(* IEC 61131-3 sources: sis-interlock-demo/src/POUs/Sis/F_VoteArchRequired, 2 files *)

(* ---- F_VoteArchRequired.decl.st ---- *)
// Назначение: требуемое число голосов M схемы голосования по таблице 5.1; 0 — для None,
//             ForcedTrip и значений вне перечисления.
// Автор:      kr0nsch
// Версия:     0.1.0
// Документ:   docs/DESIGN.md, раздел «5.10 Вспомогательные функции голосования»
// ВНИМАНИЕ:   код демонстрационный и не предназначен для систем безопасности. Реальная ПАЗ
//             требует определения SIL, сертифицированных аппаратных и программных средств
//             и валидации по ГОСТ Р МЭК 61511.
FUNCTION F_VoteArchRequired : UINT
VAR_INPUT
    eArch : E_VoteArch;   // схема голосования
END_VAR

(* ---- F_VoteArchRequired.impl.st ---- *)
CASE eArch OF
    E_VoteArch.Vote1oo1, E_VoteArch.Vote1oo2:
        F_VoteArchRequired := 1;
    E_VoteArch.Vote2oo2, E_VoteArch.Vote2oo3:
        F_VoteArchRequired := 2;
ELSE
    // None, ForcedTrip и значения вне перечисления — схемы нет
    F_VoteArchRequired := 0;
END_CASE
